// TIA Portal V21 export
// export: Created 2026-08-21T20:18:57.5210216Z, ExportSetting None, DisplayName Totally Integrated Automation Portal, DisplayVersion V21, DisplayName STEP 7 Professional, DisplayVersion V21, DisplayName STEP 7 Safety, DisplayVersion V21, DisplayName Tech WebApplication, DisplayVersion V21, DisplayName WinCC Basic/Comfort/Advanced, DisplayVersion V21, DisplayName WinCC Professional, DisplayVersion V21, DisplayName WinCC Unified, DisplayVersion V21
TYPE "UDT_Service_ConfigParaIndexType"
   STRUCT
      IndexAnalog { S7_SetPoint := 'True'} : DWord;   // Reference for Index number of the analog parameter
      IndexDigital { S7_SetPoint := 'True'} : DWord;   // Reference for Index number of the digital parameter
      IndexBinary { S7_SetPoint := 'True'} : DWord;   // Reference for Index number of the binary parameter
      IndexString { S7_SetPoint := 'True'} : DWord;   // Reference for Index number of the string parameter
   END_STRUCT;
END_TYPE
